Fanuc KAREL source: kb00065.KL

PROGRAM KB00065
%STACKSIZE=65535
%PRIORITY=65535
%NOLOCKGROUP
VAR
P1 : STRING[80]
P2 : INTEGER
P3 : INTEGER
P4 : STRING[80]
P5 : STRING[80]
P6 : INTEGER
P7 : INTEGER
P8 : INTEGER
BEGIN
P1='A'
P2=1
P3=1
P4='A'
P5='A'
P6=1
P7=1
P8=1
DISCTRL_ALPH(P1,P2,P3,P4,P5,P6,P7,P8)
END KB00065
